// TIA Portal V17 export
// export: Created 2026-11-10T15:00:48.6641979Z, ExportSetting WithDefaults, DisplayName Totally Integrated Automation Portal, DisplayVersion V17, DisplayName TIA Portal Openness, DisplayVersion V17, DisplayName TIA Portal Version Control Interface, DisplayVersion V17, DisplayName STEP 7 Professional, DisplayVersion V17, DisplayName STEP 7 Safety, DisplayVersion V17, DisplayName WinCC Advanced, DisplayVersion V17
GraphicList "Level100"  ListRange=Decimal, Mode=Simple
  GraphicListEntry   EntryType=Range, To=9, Picture=Tank_0
  GraphicListEntry   EntryType=Range, From=10, To=19, Picture=Tank_1
  GraphicListEntry   EntryType=Range, From=20, To=29, Picture=Tank_2
  GraphicListEntry   EntryType=Range, From=30, To=39, Picture=Tank_3
  GraphicListEntry   EntryType=Range, From=40, To=49, Picture=Tank_4
  GraphicListEntry   EntryType=Range, From=50, To=59, Picture=Tank_5
  GraphicListEntry   EntryType=Range, From=60, To=69, Picture=Tank_6
  GraphicListEntry   EntryType=Range, From=70, To=79, Picture=Tank_7
  GraphicListEntry   EntryType=Range, From=80, To=89, Picture=Tank_8
  GraphicListEntry   EntryType=Range, From=90, To=99, Picture=Tank_9
  GraphicListEntry   EntryType=Range, From=100, To=100, Picture=Tank_10
